# EPICS autosave request: 1.5.0/debian-12/7.0.10/modules/ADCore-ee039d2/db/NDROIStat_settings.req
$(P)$(R)TSNumPoints
$(P)$(R)TSRead.SCAN
file "NDPluginBase_settings.req", P=$(P), R=$(R)
